// TIA Portal V21 export
DATA_BLOCK "IDB_SclTimersParam"   // DB19
// stored: InstanceOfName FB_SclTimers, InstanceOfType FB
"FB_SclTimers"
   // VAR_INPUT
   //    Start : Bool;
   //    Reset : Bool;
   //    DelayTime : Time;
   // END_VAR
   // VAR_OUTPUT
   //    DelayedOn : Bool;
   //    RunOn : Bool;
   //    Pulse : Bool;
   //    Count : Int;
   //    CountReached : Bool;
   // END_VAR
   // VAR
   //    OnDelay { S7_SetPoint := 'True'} : TON_TIME;
   //    OffDelay { S7_SetPoint := 'True'} : TOF_TIME;
   //    PulseTimer { S7_SetPoint := 'True'} : TP_TIME;
   //    StartEdge { S7_SetPoint := 'True'} : R_TRIG;
   //    StopEdge { S7_SetPoint := 'True'} : F_TRIG;
   //    PartCounter { S7_SetPoint := 'True'} : CTU_INT;
   // END_VAR
BEGIN
END_DATA_BLOCK
